Staubli VAL3: MoveL.pgx

public program MoveL(pointRx x_pPoint, tool x_tTool, mdesc x_mSpeed, num& x_nMoveId, bool x_bExact)
// // 直线运动movel程序
// // 用该程序替代原val3程序中的movel()指令即可
// // 因为原move指令有返回值moveID，所以这里引入一个x_nMoveId，随参考传递出来
begin
  // ---------------------------------------------------------------------------- //
  // 直线运动movel程序
  // 用该程序替代原val3程序中的movel()指令即可
  // 因为原move指令有返回值moveID，所以这里引入一个x_nMoveId，随参考传递出来
  // ---------------------------------------------------------------------------- //
  //
  //
  //
  // 2023.03.15 pointToJoint()时，l_jRef应该取当前指令的前一个点而不是herej()，否则l_jResult可能出现错的解
  // 解决方法：1.新开一个任务，监控当前moveid，当监控开始执行该点轨迹时，重新pointToJoint()，得到l_jResult（待更新）
  x_nMoveId=movel(x_pPoint,x_tTool,x_mSpeed)
  if x_bExact
    //判断是否精确到达
    waitEndMove()
  endIf
  // log
  call logMoveMsgL(x_pPoint,x_tTool,x_mSpeed,x_nMoveId,x_bExact)

end
